Fanuc KAREL source: kt00494.KL

-- PROVISIONAL review KL for V770-1; original PC SHA256 8313a63e70eec7ee513d6d27d155825665f1a4ba4bd2f451bd9447c9f28f7cb5
-- Incomplete behavior may be omitted. Consult companion uncertainty JSON. Do not deploy.
PROGRAM KT00494
%NOLOCKGROUP
-- UNRESOLVED_DECL P1 type=000102
-- UNRESOLVED_DECL P2 type=000101
-- UNRESOLVED_DECL OUT type=000101
BEGIN
  -- UNRESOLVED_PC offsets 5-20; opcodes 2E,22,32,35
  -- UNRESOLVED_PC offsets 25-54; opcodes 49,7E,49,60,4A
  -- UNRESOLVED_PC offsets 59-63; opcodes 7F
END KT00494
